(* PLC project Claude1.project, CODESYS CODESYS V3.5 SP20 *)
(* stored: creationDateTime 2026-10-15T18:33:43.8009957, modificationDateTime 2026-10-15T18:16:57.2099678 *)

PROGRAM PLC_PRG
  VAR_INPUT
    i_bStart : BOOL;
    i_bStop : BOOL;  (* Contato NF: FALSE = emergencia acionada *)
    i_wTempSensor : INT;  (* Sinal bruto 0..27648 *)
  END_VAR
  VAR_OUTPUT
    o_bHeater : BOOL;
    o_bMixer : BOOL;
    o_rAvgTemp : REAL;
  END_VAR
  VAR
    aTempHist : ARRAY[0..4] OF REAL;
    tmrMix : TON;
    iState : INT := 0;
    iIdx : INT;
    rTempScaled : REAL;
    rSum : REAL;
    bTmrEnable : BOOL;
  END_VAR

                    
(* ===== 1. ESCALONAMENTO: 0..27648 -> 0.0..150.0 degC ===== *)
rTempScaled := (INT_TO_REAL(i_wTempSensor) * 150.0) / 27648.0;

IF rTempScaled < 0.0 THEN
    rTempScaled := 0.0;
ELSIF rTempScaled > 150.0 THEN
    rTempScaled := 150.0;
END_IF;

(* ===== 2. MEDIA MOVEL (FOR) ===== *)
FOR iIdx := 4 TO 1 BY -1 DO
    aTempHist[iIdx] := aTempHist[iIdx - 1];
END_FOR;
aTempHist[0] := rTempScaled;

rSum := 0.0;
FOR iIdx := 0 TO 4 DO
    rSum := rSum + aTempHist[iIdx];
END_FOR;
o_rAvgTemp := rSum / 5.0;

(* ===== 4. SEGURANCA E INTERLOCKS (antes da maquina de estados) ===== *)
IF NOT i_bStop THEN
    (* Emergencia acionada: estado seguro *)
    iState     := 0;
    bTmrEnable := FALSE;
    tmrMix(IN := FALSE, PT := T#10s);
    o_bHeater  := FALSE;
    o_bMixer   := FALSE;
ELSE
    (* ===== 3. MAQUINA DE ESTADOS ===== *)
    CASE iState OF

        0: (* IDLE *)
            o_bHeater  := FALSE;
            o_bMixer   := FALSE;
            bTmrEnable := FALSE;
            IF i_bStart THEN
                iState := 1;
            END_IF;

        1: (* HEATING *)
            o_bHeater := TRUE;
            o_bMixer  := FALSE;
            IF o_rAvgTemp > 80.0 THEN
                o_bHeater  := FALSE;
                o_bMixer   := TRUE;
                bTmrEnable := TRUE;
                iState     := 2;
            END_IF;

        2: (* MIXING *)
            o_bHeater := FALSE;
            o_bMixer  := TRUE;
            IF tmrMix.Q THEN
                o_bMixer   := FALSE;
                bTmrEnable := FALSE;
                iState     := 0;
            END_IF;

    ELSE
        (* Estado invalido: retorna ao estado seguro *)
        o_bHeater  := FALSE;
        o_bMixer   := FALSE;
        bTmrEnable := FALSE;
        iState     := 0;
    END_CASE;

    (* Chamada do temporizador apos a avaliacao dos estados *)
    tmrMix(IN := bTmrEnable, PT := T#10s);
END_IF;

                  
END_PROGRAM

CONFIGURATION Device
  RESOURCE Application ON PLC
    TASK MainTask(INTERVAL := T#20ms, PRIORITY := 1);
    PROGRAM PLC_PRG WITH MainTask : PLC_PRG;
  END_RESOURCE
END_CONFIGURATION
